// TIA Portal V20 export
DATA_BLOCK "DB_SYSTEM"   // DB12
{ S7_Optimized_Access := 'TRUE' }
// stored: MemoryReserve 100
   VAR RETAIN
      OP2 : Struct
         M1 { S7_SetPoint := 'True'} : Time;
         M2 { S7_SetPoint := 'True'} : Time;
         M3 { S7_SetPoint := 'True'} : Time;
         M4 { S7_SetPoint := 'True'} : Time;
         M5 { S7_SetPoint := 'True'} : Time;
         M6 { S7_SetPoint := 'True'} : Time;
         M7 { S7_SetPoint := 'True'} : Time;
         M8 { S7_SetPoint := 'True'} : Time;
      END_STRUCT;
      OP3 : Struct
         M1 { S7_SetPoint := 'True'} : Time;
         M2 { S7_SetPoint := 'True'} : Time;
         M3 { S7_SetPoint := 'True'} : Time;
         M4 { S7_SetPoint := 'True'} : Time;
         M5 { S7_SetPoint := 'True'} : Time;
         M6 { S7_SetPoint := 'True'} : Time;
         M7 { S7_SetPoint := 'True'} : Time;
         M8 { S7_SetPoint := 'True'} : Time;
      END_STRUCT;
   END_VAR
BEGIN
END_DATA_BLOCK
